(* IEC 61131-3 sources: PortalRobot/Portal_robot/Device/application/ST/ST_MACHINE, 19 files *)

(* ---- E_MACHINE_OPERATION.st ---- *)
{attribute 'qualified_only'}
{attribute 'strict'}
TYPE E_MACHINE_OPERATION :
(
	NONE,
    LOAD,
    UNLOAD,
    CHANGE
);
END_TYPE

(* ---- E_MACHINE_POINTS.st ---- *)
{attribute 'qualified_only'}
{attribute 'strict'}
TYPE E_MACHINE_POINTS :
(
	NONE,
	ABOVE,
    INSIDE,
    CHUCK_APPROACH,
    CHUCK
);
END_TYPE

(* ---- E_MACHINE_STATE.st ---- *)
{attribute 'qualified_only'}
{attribute 'strict'}
TYPE E_MACHINE_STATE :
(
	DISABLED := 0,
	OPERATOR_CHOICE_PART,
	OPERATOR_CHOICE_RUN,
	OPERATOR_CHOICE_DOOR,
    IDLE,
	CHOSE,
	READ,
	NEXT,
	RELEASE_ROBOT_ACTION,
	ROBOT_MOVE,
	ROBOT_ACTION,
	DOOR_OPEN,
	DOOR_CLOSE,
	CHUCK_OPEN,
	CHUCK_CLOSE,
	CYCLE_START,
	DONE,
	ERROR
);
END_TYPE

(* ---- E_PART_STATE.st ---- *)
{attribute 'qualified_only'}
{attribute 'strict'}
TYPE E_PART_STATE :
(
	UNKNOWN := 0,
    EMPTY   := 1,
    LOADED  := 2
);
END_TYPE

(* ---- E_PART_TYPE.st ---- *)
{attribute 'qualified_only'}
{attribute 'strict'}
TYPE E_PART_TYPE :
(
	UNKNOWN,
	DETAIL,
	PART
);
END_TYPE

(* ---- ST_MACHINE_COMMAND.st ---- *)
TYPE ST_MACHINE_COMMAND :
STRUCT
	stIo    : ST_MACHINE_IO_COMMAND; // Команды исполнительным механизмам станка
	stRobot : ST_ROBOT_COMMAND; // Команда роботу от алгоритма станка
END_STRUCT
END_TYPE

(* ---- ST_MACHINE_DIAG.st ---- *)
TYPE ST_MACHINE_DIAG :
STRUCT
	eState            : E_MACHINE_STATE; // Текущее состояние автомата станка
	eGrantedOperation : E_MACHINE_OPERATION; // Разрешённая операция
	eActualOperation  : E_MACHINE_OPERATION; // Выполняемая операция
	stWarning         : ST_WARNING_EVENT; // Последнее предупреждение станка
END_STRUCT
END_TYPE

(* ---- ST_MACHINE_ERROR.st ---- *)
TYPE ST_MACHINE_ERROR :
STRUCT
	WRONG_OPERATION : BOOL; // Не удалось выбрать операцию
	WRONG_COMMAND   : BOOL; // В рецепте встретилась неизвестная команда
	ROBOT_MOTION    : BOOL; // Ошибка перемещения робота
	ROBOT_ACTION    : BOOL; // Ошибка действия захвата
	DOOR_OPEN       : BOOL; // Не удалось открыть дверь
	DOOR_CLOSE      : BOOL; // Не удалось закрыть дверь
	CHUCK_OPEN      : BOOL; // Не удалось разжать патрон
	CHUCK_CLOSE     : BOOL; // Не удалось зажать патрон
	CYCLE_START     : BOOL; // Не удалось запустить цикл станка
	SAFETY_STOP     : BOOL; // Получена глобальная ошибка ячейки
	UNKNOWN_DETAIL  : BOOL; // Неизвестно состояние детали в станке
	MACHINE_ALARM   : BOOL; // Станок сообщил аварию
	INDEX_ERROR     : BOOL; // Индекс рецепта вышел за границы
	DOOR_ROBOT      : BOOL; // Дверь закрыта при нахождении робота внутри
	MACHINE_IDLE    : BOOL; // Авария станка возникла в ожидании
	TIMEOUT_ROBOT_MOVE    : BOOL; // Превышено время перемещения робота
	TIMEOUT_ROBOT_ACTION  : BOOL; // Превышено время действия захвата
	TIMEOUT_ROBOT_RELEASE : BOOL; // Робот не освободил интерфейс команды вовремя
	TIMEOUT_DOOR_OPEN     : BOOL; // Превышено время открытия двери
	TIMEOUT_DOOR_CLOSE    : BOOL; // Превышено время закрытия двери
	TIMEOUT_HATCH_UNLOCK  : BOOL; // Превышено время открытия замка роботного люка
	TIMEOUT_CHUCK_OPEN    : BOOL; // Превышено время разжима патрона
	TIMEOUT_CHUCK_CLOSE   : BOOL; // Превышено время зажима патрона
	TIMEOUT_CYCLE_START   : BOOL; // Превышено время подтверждения запуска цикла
	SAFETY_DOOR_OPEN     : BOOL; // Операторская дверь открылась во время обслуживания
	HATCH_UNLOCK_PROCESSING : BOOL; // Замок открыт во время обработки в автоматической линии
END_STRUCT
END_TYPE

(* ---- ST_MACHINE_ERRORS.st ---- *)
TYPE ST_MACHINE_ERRORS :
STRUCT
	dwErrorActive : DWORD; // Битовая маска активных ошибок
	dwErrorLast   : DWORD; // Битовая маска последних ошибок
	dwAlarmActive : DWORD; // Собственные аварии станка для общего журнала
	stErrorActive : ST_MACHINE_ERROR; // Расшифровка активных ошибок
	stErrorLast   : ST_MACHINE_ERROR; // Расшифровка последних ошибок
END_STRUCT
END_TYPE

(* ---- ST_MACHINE_FAULT_REQUEST.st ---- *)
TYPE ST_MACHINE_FAULT_REQUEST :
STRUCT
	xEnabled             : BOOL; // Глобальное разрешение диагностической инъекции
	xReset               : BOOL; // Отдельный сброс источника неисправности станка
	xMachineAlarm        : BOOL; // Общая авария виртуального станка
	xDoorFault           : BOOL; // Неисправность механизма двери
	xChuckFault          : BOOL; // Неисправность механизма патрона
	xTimeoutRobotMove    : BOOL; // Не подтверждать завершение движения робота
	xTimeoutRobotAction  : BOOL; // Не подтверждать действие захвата
	xTimeoutRobotRelease : BOOL; // Не подтверждать освобождение интерфейса робота
	xTimeoutDoorOpen     : BOOL; // Не подтверждать открытие двери
	xTimeoutDoorClose    : BOOL; // Не подтверждать закрытие двери
	xTimeoutHatchUnlock  : BOOL; // Не подтверждать открытие замка до TIMEOUT
	xTimeoutChuckOpen    : BOOL; // Не подтверждать разжим патрона
	xTimeoutChuckClose   : BOOL; // Не подтверждать зажим патрона
	xTimeoutCycleStart   : BOOL; // Не подтверждать запуск цикла обработки
END_STRUCT
END_TYPE

(* ---- ST_MACHINE_IO_COMMAND.st ---- *)
TYPE ST_MACHINE_IO_COMMAND :
STRUCT
	xOpenDoor       : BOOL; // Открыть роботный люк; имя сохранено для совместимости
	xCloseDoor      : BOOL; // Закрыть роботный люк; имя сохранено для совместимости
	xHatchUnLock    : BOOL; // Открыть замок роботного люка; FALSE удерживает замок закрытым
	xOpenSafetyDoor : BOOL; // Открыть операторскую дверь
	xCloseSafetyDoor: BOOL; // Закрыть операторскую дверь
	xClampChuck   : BOOL; // Зажать патрон
	xUnclampChuck : BOOL; // Разжать патрон
	xStartCycle   : BOOL; // Запустить обработку
	xReset        : BOOL; // Сбросить аварию станка
END_STRUCT
END_TYPE

(* ---- ST_MACHINE_IO_STATUS.st ---- *)
TYPE ST_MACHINE_IO_STATUS :
STRUCT
	xReady          : BOOL; // Станок готов принимать команды
	xAlarm          : BOOL; // Активна авария станка
	xDoorOpen       : BOOL; // Роботный люк открыт; имя сохранено для совместимости
	xDoorClosed     : BOOL; // Роботный люк закрыт; имя сохранено для совместимости
	xHatchLocked    : BOOL; // Замок роботного люка закрыт (0 — открыт, 1 — закрыт)
	xSafetyDoorOpen   : BOOL; // Операторская дверь открыта
	xSafetyDoorClosed : BOOL; // Операторская дверь закрыта
	xChuckClamped   : BOOL; // Патрон зажат
	xChuckUnclamped : BOOL; // Патрон разжат
	xCycleActive    : BOOL; // Выполняется цикл обработки
	xCycleDone      : BOOL; // Цикл обработки завершён
	tRemaining      : TIME; // Оставшееся время обработки
END_STRUCT
END_TYPE

(* ---- ST_MACHINE_POINTS.st ---- *)
TYPE ST_MACHINE_POINTS :
STRUCT
	eNone          : E_POINT_NAME; // Пустое имя точки
	eAbove         : E_POINT_NAME; // Точка над рабочей зоной станка
	eInside        : E_POINT_NAME; // Точка внутри рабочей зоны станка
	eChuckApproach : E_POINT_NAME; // Точка подхода к патрону
	eChuck         : E_POINT_NAME; // Рабочая точка патрона
END_STRUCT
END_TYPE

(* ---- ST_MACHINE_PUBLIC.st ---- *)
TYPE ST_MACHINE_PUBLIC :
STRUCT
	xEnabled             : BOOL; // Станок включен в работу
	xDisablePending      : BOOL; // Запрошено отключение после выхода автомата в разрешённый шаг
	xPowerAllowed        : BOOL; // Кнопка включения, отключения или отмены отключения доступна
	xResetAllowed        : BOOL; // Кнопка сброса ошибки станка доступна
	xManualControlAllowed       : BOOL; // Ручное управление разрешено режимом и состоянием станка
	xManualSafetyDoorControlEnabled : BOOL; // Операторская дверь управляется только моделью
	xManualSafetyDoorOpenAllowed : BOOL; // Разрешено открыть операторскую дверь
	xManualSafetyDoorCloseAllowed: BOOL; // Разрешено закрыть операторскую дверь
	xManualHatchOpenAllowed      : BOOL; // Разрешено открыть роботный люк
	xManualHatchCloseAllowed     : BOOL; // Разрешено закрыть роботный люк
	xManualHatchUnlockAllowed    : BOOL; // Разрешено открыть замок роботного люка
	xManualHatchLockAllowed      : BOOL; // Разрешено закрыть замок роботного люка
	xManualChuckOpenAllowed      : BOOL; // Разрешено разжать патрон
	xManualChuckCloseAllowed     : BOOL; // Разрешено зажать патрон
	xProcessing          : BOOL; // Станок выполняет цикл обработки
    xPartReady           : BOOL; // Обработка детали завершена
    xServiceRequired     : BOOL; // Станку требуется обслуживание роботом
    xCanAcceptService    : BOOL; // Станок готов принять робота
    xRobotReleased       : BOOL; // Робот освобождён после операции
	xDone                : BOOL; // Операция обслуживания завершена
    xBusy                : BOOL; // Блок выполняет операцию обслуживания
    xError               : BOOL; // Станок находится в ошибке
	xCriticalError       : BOOL; // Ошибка требует зависимой аварии и остановки робота
	xAlarmError          : BOOL; // Активна первичная ошибка оборудования станка
	xExternalError       : BOOL; // Активна внешняя ошибка
	xServiceRejected     : BOOL; // Обслуживание безопасно отклонено до входа робота в станок
    xDoorOpen            : BOOL; // Дверь станка открыта
    xAlarm               : BOOL; // Активна авария станка
	stIo    			 : ST_MACHINE_IO_STATUS; // Статусы исполнительных механизмов станка
    eRecommendedOperation: E_MACHINE_OPERATION; // Рекомендуемая операция обслуживания
    ePartState           : E_PART_STATE; // Состояние детали в патроне
    ePartType            : E_PART_TYPE; // Тип изделия в патроне: заготовка или готовая деталь
    eAbovePoint          : E_POINT_NAME; // Имя точки над станком
    lrAboveX             : LREAL; // Координата X точки над станком
	tCycleExpected       : TIME; // Ожидаемое время текущего цикла
	tCycleElapsed        : TIME; // Прошедшее время текущего цикла
	tMeasuredCycle       : TIME; // Последнее измеренное время корректного автоцикла
	tRemaining           : TIME; // Оставшееся время обработки
	xCycleTimeValid      : BOOL; // Доступна оценка времени цикла
	xMeasuredTimeValid   : BOOL; // Получено измерение корректного автоцикла
	xCycleOvertime       : BOOL; // Фактический цикл превысил ожидаемое время
END_STRUCT
END_TYPE

(* ---- ST_MACHINE_RECIPE.st ---- *)
TYPE ST_MACHINE_RECIPE :
STRUCT
	eRobotAction    : E_ROBOT_ACTION; // Действие робота на шаге рецепта
	eCommand        : E_MACHINE_STATE; // Команда шага рецепта
	stPoint         : E_MACHINE_POINTS; // Логическая точка станка
	xRetreatStarted : BOOL; // Признак начала отхода робота
	xRobotDone      : BOOL; // Признак освобождения робота после шага
END_STRUCT
END_TYPE

(* ---- ST_MACHINE_SIM_DIAG.st ---- *)
TYPE ST_MACHINE_SIM_DIAG :
STRUCT
	xDoorOpening   : BOOL; // Выполняется открытие роботного люка
	xDoorClosing   : BOOL; // Выполняется закрытие роботного люка
	xSafetyDoorOpening : BOOL; // Выполняется открытие операторской двери
	xSafetyDoorClosing : BOOL; // Выполняется закрытие операторской двери
	xChuckClamping : BOOL; // Выполняется зажим патрона
	xChuckOpening  : BOOL; // Выполняется разжим патрона
	xCycleStarting : BOOL; // Выполняется запуск цикла
	xResetAllowed  : BOOL; // Источник имитации снят и авария симулятора может быть сброшена
END_STRUCT
END_TYPE

(* ---- ST_MACHINE_SIM_ERROR.st ---- *)
TYPE ST_MACHINE_SIM_ERROR :
STRUCT
	MACHINE_ALARM : BOOL; // Активна имитация аварии станка
	DOOR_FAULT    : BOOL; // Ошибка механизма двери
	CHUCK_FAULT   : BOOL; // Ошибка механизма патрона
END_STRUCT
END_TYPE

(* ---- ST_MACHINE_SIM_ERRORS.st ---- *)
TYPE ST_MACHINE_SIM_ERRORS :
STRUCT
	dwErrorActive : DWORD; // Битовая маска активных ошибок
	dwErrorLast   : DWORD; // Битовая маска последних ошибок
	stErrorActive : ST_MACHINE_SIM_ERROR; // Расшифровка активных ошибок
	stErrorLast   : ST_MACHINE_SIM_ERROR; // Расшифровка последних ошибок
END_STRUCT
END_TYPE

(* ---- ST_MACHINE_TIMEOUTS.st ---- *)
TYPE ST_MACHINE_TIMEOUTS :
STRUCT
	tRobotMove    : TIME := T#60S; // Допустимое время движения робота
	tRobotAction  : TIME := T#10S; // Допустимое время действия захвата
	tRobotRelease : TIME := T#5S; // Допустимое время освобождения интерфейса робота
	tDoorOpen     : TIME := T#10S; // Допустимое время открытия двери
	tDoorClose    : TIME := T#10S; // Допустимое время закрытия двери
	tHatchUnlock  : TIME := T#5S; // Допустимое ожидание открытия замка роботного люка
	tChuckOpen    : TIME := T#10S; // Допустимое время разжима патрона
	tChuckClose   : TIME := T#10S; // Допустимое время зажима патрона
	tCycleStart   : TIME := T#10S; // Допустимое время подтверждения запуска цикла
END_STRUCT
END_TYPE
